{attribute 'qualified_only'}
//{attribute 'strict'}
{attribute 'to_string'}
TYPE E_CIP_Usage :
(
	eNotInUse := 0,
	eTank_1,
	eTank_2,
	eTank_3,
	eTank_4,
	eTriBlender_Marinada,
	eTriBlender_Color,
	eLine_Marinada,
	eLine_Color,
	eLocal,
	eExternal	//GAD client through Siemens, stays after eLocal: arr_CIP_Param ends at eLocal
	//,eClient
);
END_TYPE

(* stored: Version 1.1.0.1, ProductVersion 3.1.4024.12
   DUT E_CIP_Usage: Id {62ed165f-f4bd-4351-99d8-f631457fb546} *)
